Fanuc KAREL source: KT00661.KL

PROGRAM KT00661
%NOLOCKGROUP
VAR
  P1: XYZWPR
  P2: XYZWPR
  OUT: INTEGER
BEGIN
  P1.X = 1.0
  P2.Y = 2.0
  P1.X = 1.0
  P2.Y = 2.0
  OUT = NOT P1
END KT00661
